FUNCTION F_Double (* Verdoppelt einen INT-Wert *)
  (* Standard: 61499-1; Description: Copyright (c) 2026 Meisterschulen am Ostbahnhof This program and the accompanying materials are made available under the terms of the Eclipse Public License 2.0 which is available at https://www.eclipse.org/legal/epl-2.0/ SPDX-License-Identifier: EPL-2.0 *)
  (* Version 1.0, 2026-10-16, Franz Höpfinger, Meisterschulen am Ostbahnhof, Uebung: Function in ST aus GCF/FB aufrufen *)
  PACKAGE Meins::GcfFunctionCall;
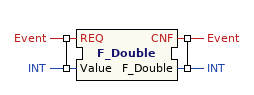
  EVENT_INPUT
    REQ WITH Value;
  END_EVENT
  EVENT_OUTPUT
    CNF WITH F_Double;
  END_EVENT
  VAR_INPUT
    Value : INT;
  END_VAR
  VAR_OUTPUT
    F_Double : INT;
  END_VAR
  BODY IN ST:
PACKAGE Meins::GcfFunctionCall;

(* Verdoppelt einen INT-Wert *)
FUNCTION F_Double : INT

VAR_INPUT
	Value : INT;
END_VAR

F_Double := Value * 2;

END_FUNCTION
  END_BODY
END_FUNCTION
